FUNCTION F_ConvArrBitsToWord_1 : WORD
VAR_INPUT
	arrBits: ARRAY [0..15] OF BOOL;
END_VAR
VAR
END_VAR

F_ConvArrBitsToWord := 0;

END_FUNCTION

(* stored: Version 1.1.0.1, ProductVersion 3.1.4024.15
   POU F_ConvArrBitsToWord_1: Id {57f351d0-4170-4314-9b0a-4542dea5b017}, SpecialFunc None *)
